// TIA Portal V21 export
DATA_BLOCK "IDB_AnaTimerInIf"   // DB8
// stored: InstanceOfName FB_AnaTimerInIf, InstanceOfType FB
"FB_AnaTimerInIf"
   // VAR_INPUT
   //    Enable : Bool;
   //    Start : Bool;
   // END_VAR
   // VAR_OUTPUT
   //    Done : Bool;
   // END_VAR
   // VAR
   //    Delay { S7_SetPoint := 'True'} : TON_TIME;
   // END_VAR
BEGIN
END_DATA_BLOCK
